(* Logix 5000 project; controller CIP_14485201 vendor 1 type 14 code 216 rev 38.11; software revision 38.01; part 10 of 11 *)
(* tags used below, declared in another part *)
   Bit : BOOL[128];   // BIT
   CIP_to_Process : CIP_to_Process;   // CIP TO PROCESS SIGNALS
   cipToProcess : BOOL;   // send signal to dcs
   Heartbeat_to_dcs_off : TIMER;   // 5 second toggle
   heartbeat_to_dcs_on : TIMER;   // turns on heartbeat to dcs
   Messages_List : STRING;   // ACTIVE MESSAGES ECHO FROM HMI
   MOA_Drain_Flow_Mod_Value : INT;   // PV MOA DRAIN FLOW MODULATION VALUE
   MOA_Drain_Flow_Mod_Value_Status : BOOL;   // PV MOA DRAIN FLOW MODULATION VALUE STATUS BIT
   MOA_OFF : DINT[20];   // PANELVIEW MOA OFF
   MOA_ON : DINT[20];   // PANELVIEW MOA ON
   Opcode_Description : STRING;   // ACTIVE OPCODE ECHO FROM HMI
   OpCode_Pin : DINT[5];   // OPCODE PIN ARRAY
   Panelview : INT[40];   // PANELVIEW CONTROL
   PID2 : PID;   // SUPPLY FLOW PID
   Process_Heartbeat_Memory : BOOL;
   Process_to_CIP : Process_to_CIP;   // PROCESS SIGNALS TO CIP
   pv_step_time_minutes : DINT;   // PANELVIEW DISPLAY STEP TIME MINUTES
   pv_step_time_seconds : DINT;   // PANELVIEW DISPLAY STEP TIME SECONDS
   Recipe : RECIPE[41];   // RECIPES
   SCLD_Drain_Flow : SCALE;   // DRAIN FLOW MODULATION 0-100%
   SCLD_DrainValve_Feedback : SCALE;   // DRAIN FLOW FEEDBACK POSITION 0-100%
   SCLD_Return_Temp : SCALE;   // RETURN TEMPERATURE 0-100°C
   SCLD_Rinse_Cond : SCALE;   // RINSE CONDUCTIVITY 0-10 uS/cm
   SCLD_Supply_Flow : SCALE;   // SUPPLY FLOW 0-60 GPM
   SCLD_Supply_Press : SCALE;   // SUPPLY PRESSURE 0-100 PSIG
   SCLD_Supply_Temp : SCALE;   // SUPPLY TEMPERATURE 0-100°C
   SCLD_SupplyValve_Feedback : SCALE;   // SUPPLY FLOW FEEDBACK POSITION 0-100%
   SCLD_Wash_Cond : SCALE;   // WASH CONDUCTIVITY 0-100 mS/cm
   Sequencer : CONTROL[4];   // SEQUENCER
   SP_Drain_Flow : REAL;   // CURRENT DRAIN FLOW MODULATION SETPOINT
   SP_DrainValve_HighDeadband : REAL;   // CURRENT DRAIN VALVE DEADBAND SETPOINT
   SP_DrainValve_LowDeadband : REAL;   // CURRENT DRAIN VALVE DEADBAND SETPOINT
   SP_Supply_Flow : REAL;   // CURRENT SUPPLY FLOW SETPOINT
   SP_SupplyValve_HighDeadband : REAL;   // CURRENT SUPPLY VALVE DEADBAND SETPOINT
   SP_SupplyValve_LowDeadband : REAL;   // CURRENT SUPPLY VALVE DEADBAND SETPOINT
   Step_Time_Min : STRING;
   Step_Time_Remaining : STRING[5];
   Step_Time_Sec : STRING;
   Timer : TIMER[99];   // TIMER
   Timer_Chem1_Pump : TIMER[7];   // CHEM #1 CONTROL TIMERS
   Timer_Chem2_Pump : TIMER[7];   // CHEM #2 CONTROL TIMERS
   Utility_Out : DINT[5];   // PANELVIEW UTILITY OUTPUT CONTROL
(* MainProgram, continued *)

ROUTINE _88_LEVEL   (* ladder *)
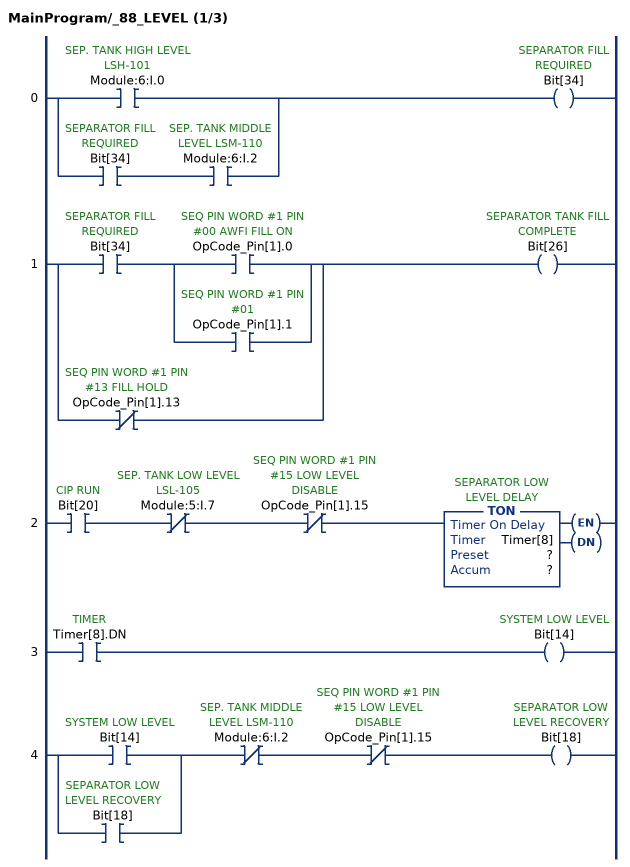
   0: [XIC(Module:6:I.0) ,XIC(Bit[34]) XIC(Module:6:I.2) ]OTE(Bit[34]);
   1: [XIC(Bit[34]) [XIC(OpCode_Pin[1].0) ,XIC(OpCode_Pin[1].1) ] ,XIO(OpCode_Pin[1].13) ]OTE(Bit[26]);
   2: XIC(Bit[20])XIO(Module:5:I.7)XIO(OpCode_Pin[1].15)TON(Timer[8],?,?);
   3: XIC(Timer[8].DN)OTE(Bit[14]);
   4: [XIC(Bit[14]) ,XIC(Bit[18]) ]XIO(Module:6:I.2)XIO(OpCode_Pin[1].15)OTE(Bit[18]);
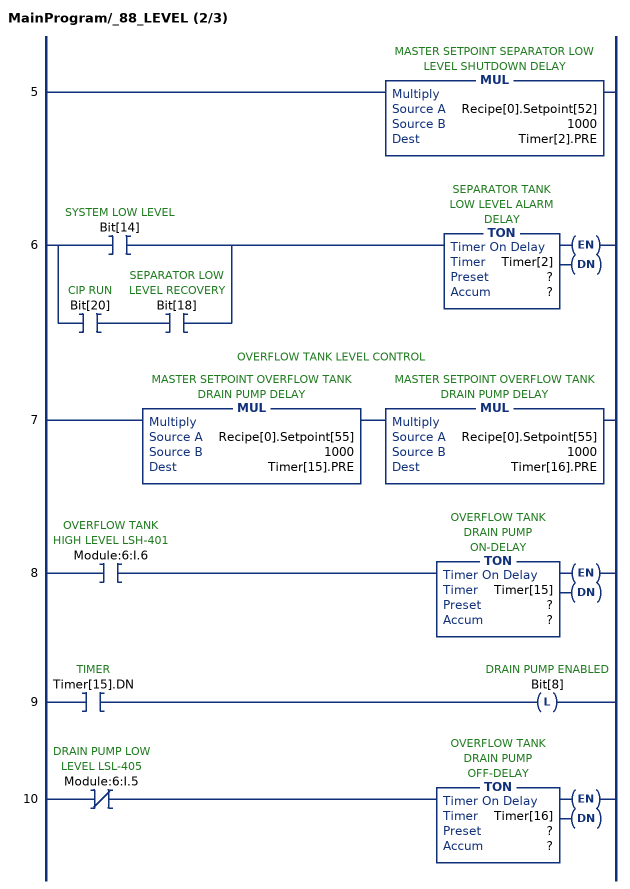
   5: MUL(Recipe[0].Setpoint[52],1000,Timer[2].PRE);
   6: [XIC(Bit[14]) ,XIC(Bit[20]) XIC(Bit[18]) ]TON(Timer[2],?,?);
   // OVERFLOW TANK LEVEL CONTROL
   7: MUL(Recipe[0].Setpoint[55],1000,Timer[15].PRE)MUL(Recipe[0].Setpoint[55],1000,Timer[16].PRE);
   8: XIC(Module:6:I.6)TON(Timer[15],?,?);
   9: XIC(Timer[15].DN)OTL(Bit[8]);
   10: XIO(Module:6:I.5)TON(Timer[16],?,?);
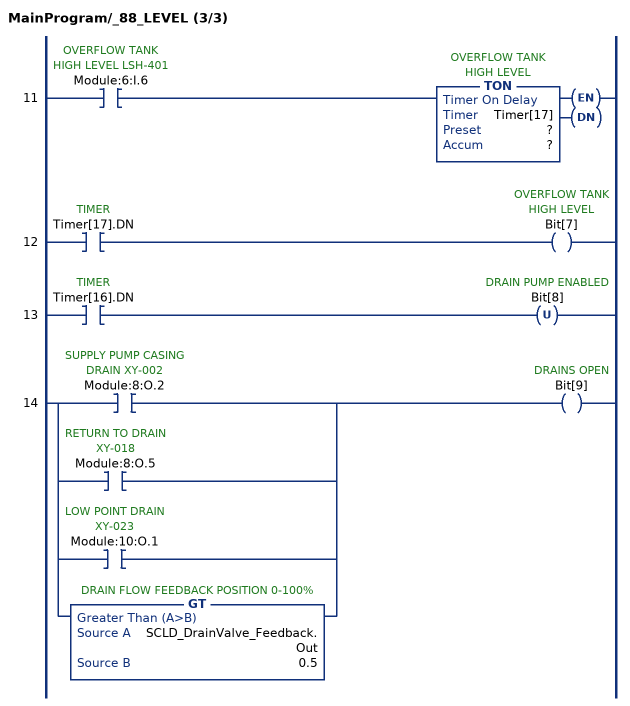
   11: XIC(Module:6:I.6)TON(Timer[17],?,?);
   12: XIC(Timer[17].DN)OTE(Bit[7]);
   13: XIC(Timer[16].DN)OTU(Bit[8]);
   14: [XIC(Module:8:O.2) ,XIC(Module:8:O.5) ,XIC(Module:10:O.1) ,GT(SCLD_DrainValve_Feedback.Out,0.5) ]OTE(Bit[9]);
END_ROUTINE

ROUTINE _89_FLOW   (* ladder *)
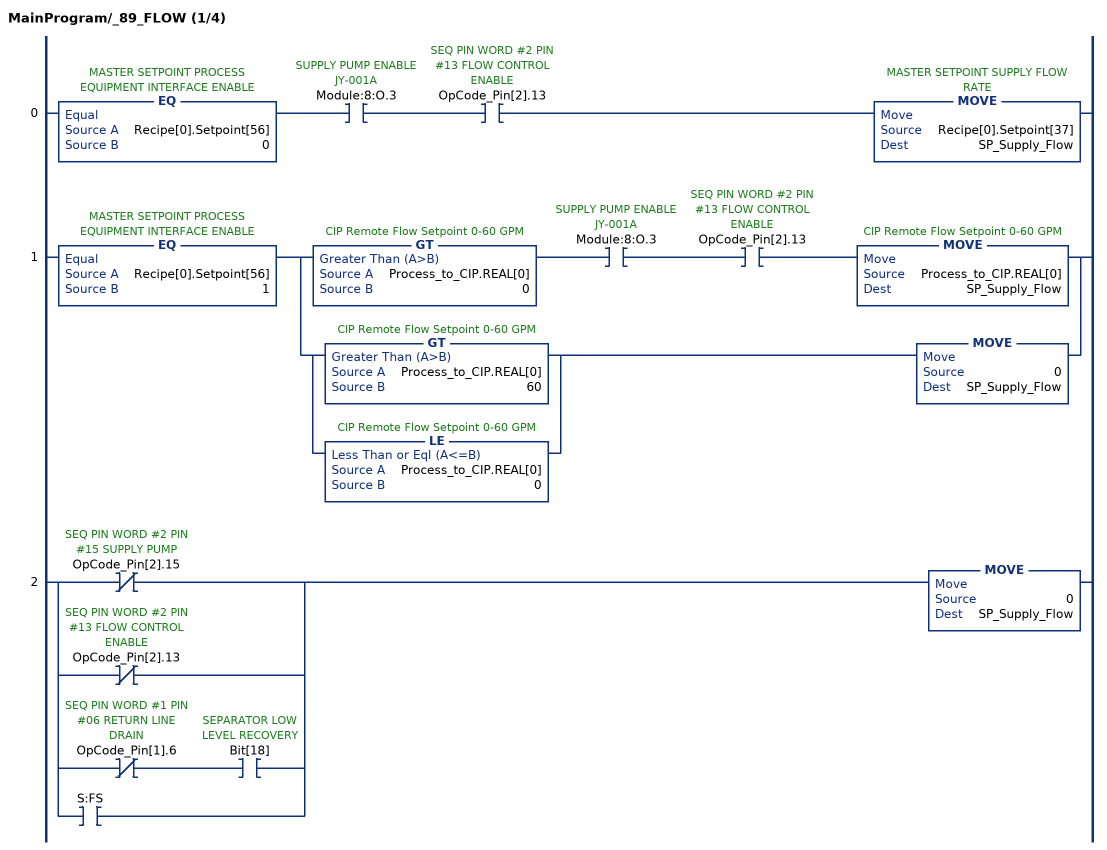
   0: EQ(Recipe[0].Setpoint[56],0)XIC(Module:8:O.3)XIC(OpCode_Pin[2].13)MOVE(Recipe[0].Setpoint[37],SP_Supply_Flow);
   1: EQ(Recipe[0].Setpoint[56],1)[GT(Process_to_CIP.REAL[0],0) XIC(Module:8:O.3) XIC(OpCode_Pin[2].13) MOVE(Process_to_CIP.REAL[0],SP_Supply_Flow) ,[GT(Process_to_CIP.REAL[0],60) ,LE(Process_to_CIP.REAL[0],0) ] MOVE(0,SP_Supply_Flow) ];
   2: [XIO(OpCode_Pin[2].15) ,XIO(OpCode_Pin[2].13) ,XIO(OpCode_Pin[1].6) XIC(Bit[18]) ,XIC(S:FS) ]MOVE(0,SP_Supply_Flow);
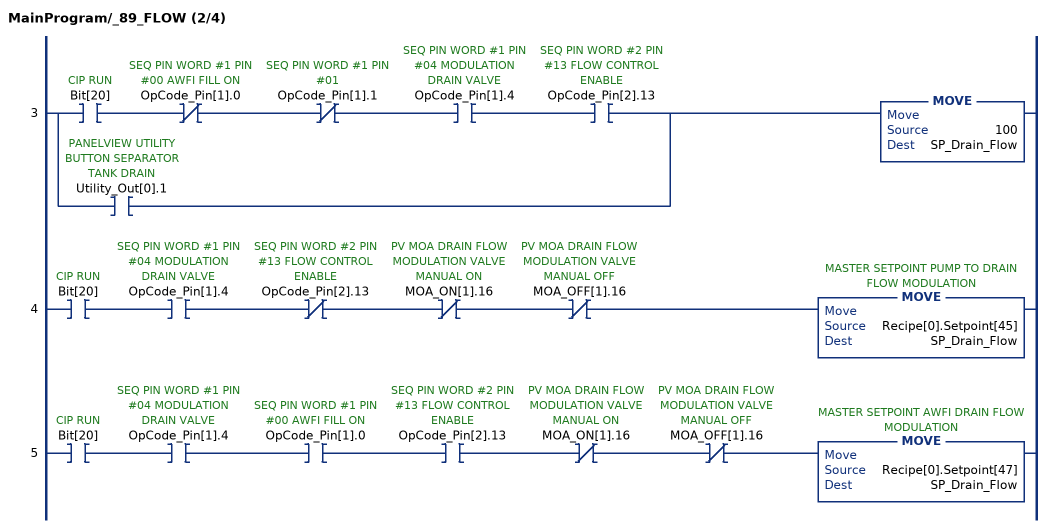
   3: [XIC(Bit[20]) XIO(OpCode_Pin[1].0) XIO(OpCode_Pin[1].1) XIC(OpCode_Pin[1].4) XIC(OpCode_Pin[2].13) ,XIC(Utility_Out[0].1) ]MOVE(100,SP_Drain_Flow);
   4: XIC(Bit[20])XIC(OpCode_Pin[1].4)XIO(OpCode_Pin[2].13)XIO(MOA_ON[1].16)XIO(MOA_OFF[1].16)MOVE(Recipe[0].Setpoint[45],SP_Drain_Flow);
   5: XIC(Bit[20])XIC(OpCode_Pin[1].4)XIC(OpCode_Pin[1].0)XIC(OpCode_Pin[2].13)XIO(MOA_ON[1].16)XIO(MOA_OFF[1].16)MOVE(Recipe[0].Setpoint[47],SP_Drain_Flow);
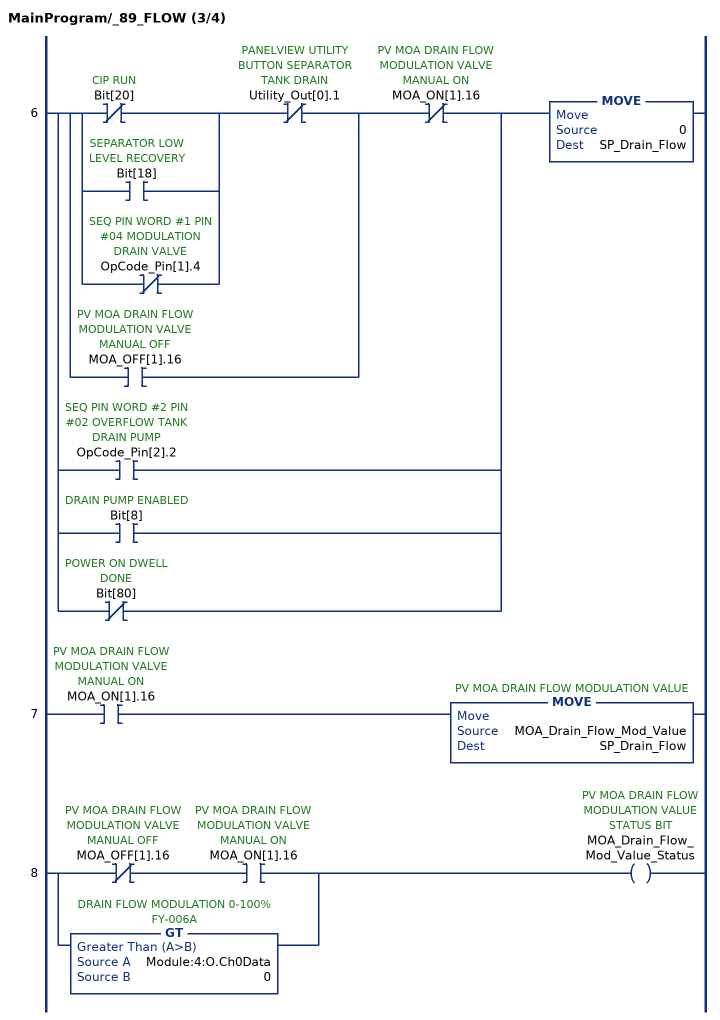
   6: [[[XIO(Bit[20]) ,XIC(Bit[18]) ,XIO(OpCode_Pin[1].4) ] XIO(Utility_Out[0].1) ,XIC(MOA_OFF[1].16) ] XIO(MOA_ON[1].16) ,XIC(OpCode_Pin[2].2) ,XIC(Bit[8]) ,XIO(Bit[80]) ]MOVE(0,SP_Drain_Flow);
   7: XIC(MOA_ON[1].16)MOVE(MOA_Drain_Flow_Mod_Value,SP_Drain_Flow);
   8: [XIO(MOA_OFF[1].16) XIC(MOA_ON[1].16) ,GT(Module:4:O.Ch0Data,0) ]OTE(MOA_Drain_Flow_Mod_Value_Status);
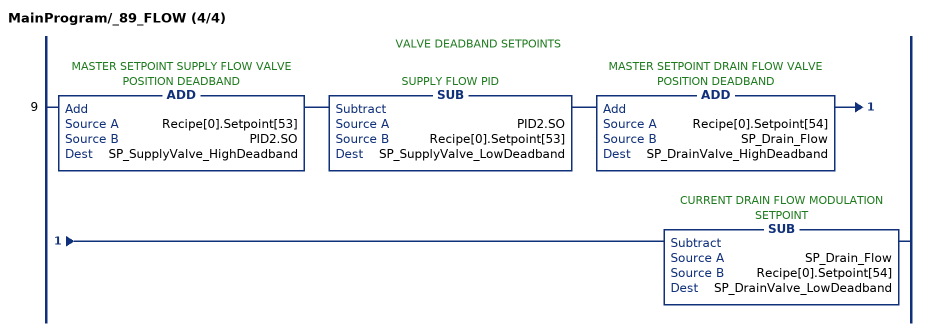
   // VALVE DEADBAND SETPOINTS
   9: ADD(Recipe[0].Setpoint[53],PID2.SO,SP_SupplyValve_HighDeadband)SUB(PID2.SO,Recipe[0].Setpoint[53],SP_SupplyValve_LowDeadband)ADD(Recipe[0].Setpoint[54],SP_Drain_Flow,SP_DrainValve_HighDeadband)SUB(SP_Drain_Flow,Recipe[0].Setpoint[54],SP_DrainValve_LowDeadband);
END_ROUTINE

ROUTINE _90_OUTPUTS   (* ladder *)
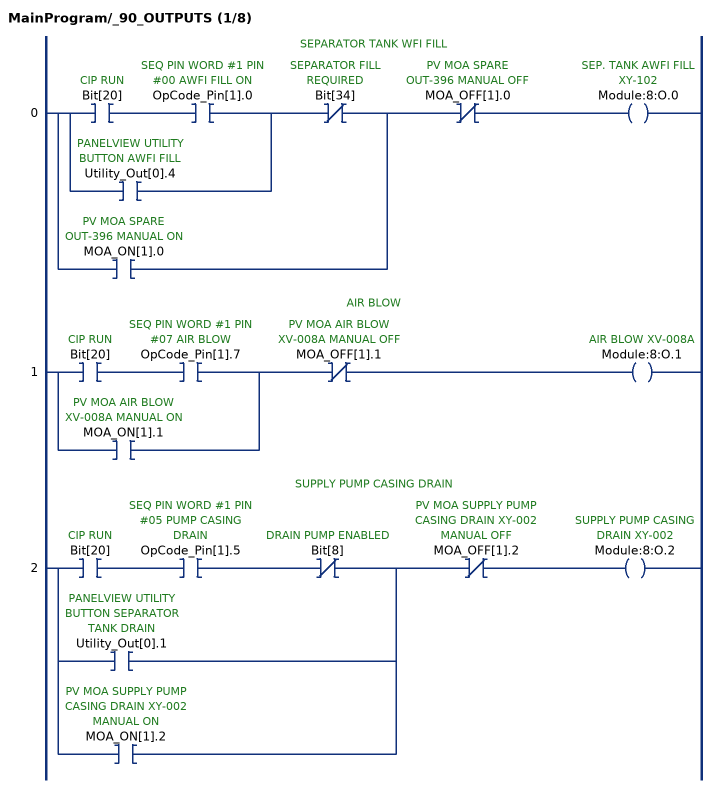
   // SEPARATOR TANK WFI FILL
   0: [[XIC(Bit[20]) XIC(OpCode_Pin[1].0) ,XIC(Utility_Out[0].4) ] XIO(Bit[34]) ,XIC(MOA_ON[1].0) ]XIO(MOA_OFF[1].0)OTE(Module:8:O.0);
   // AIR BLOW
   1: [XIC(Bit[20]) XIC(OpCode_Pin[1].7) ,XIC(MOA_ON[1].1) ]XIO(MOA_OFF[1].1)OTE(Module:8:O.1);
   // SUPPLY PUMP CASING DRAIN
   2: [XIC(Bit[20]) XIC(OpCode_Pin[1].5) XIO(Bit[8]) ,XIC(Utility_Out[0].1) ,XIC(MOA_ON[1].2) ]XIO(MOA_OFF[1].2)OTE(Module:8:O.2);
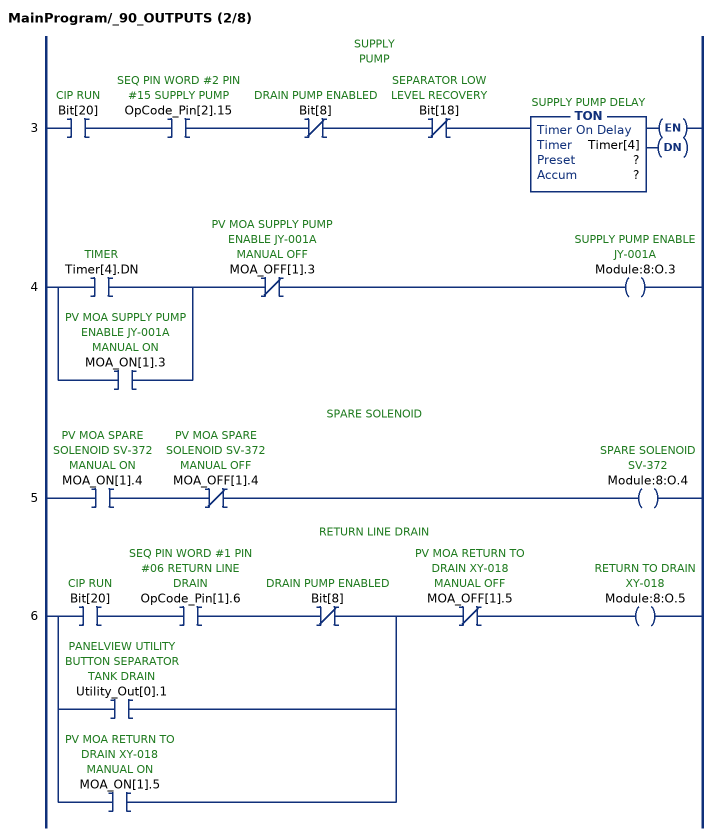
   // SUPPLY
   // PUMP
   3: XIC(Bit[20])XIC(OpCode_Pin[2].15)XIO(Bit[8])XIO(Bit[18])TON(Timer[4],?,?);
   4: [XIC(Timer[4].DN) ,XIC(MOA_ON[1].3) ]XIO(MOA_OFF[1].3)OTE(Module:8:O.3);
   // SPARE SOLENOID
   5: XIC(MOA_ON[1].4)XIO(MOA_OFF[1].4)OTE(Module:8:O.4);
   // RETURN LINE DRAIN
   6: [XIC(Bit[20]) XIC(OpCode_Pin[1].6) XIO(Bit[8]) ,XIC(Utility_Out[0].1) ,XIC(MOA_ON[1].5) ]XIO(MOA_OFF[1].5)OTE(Module:8:O.5);
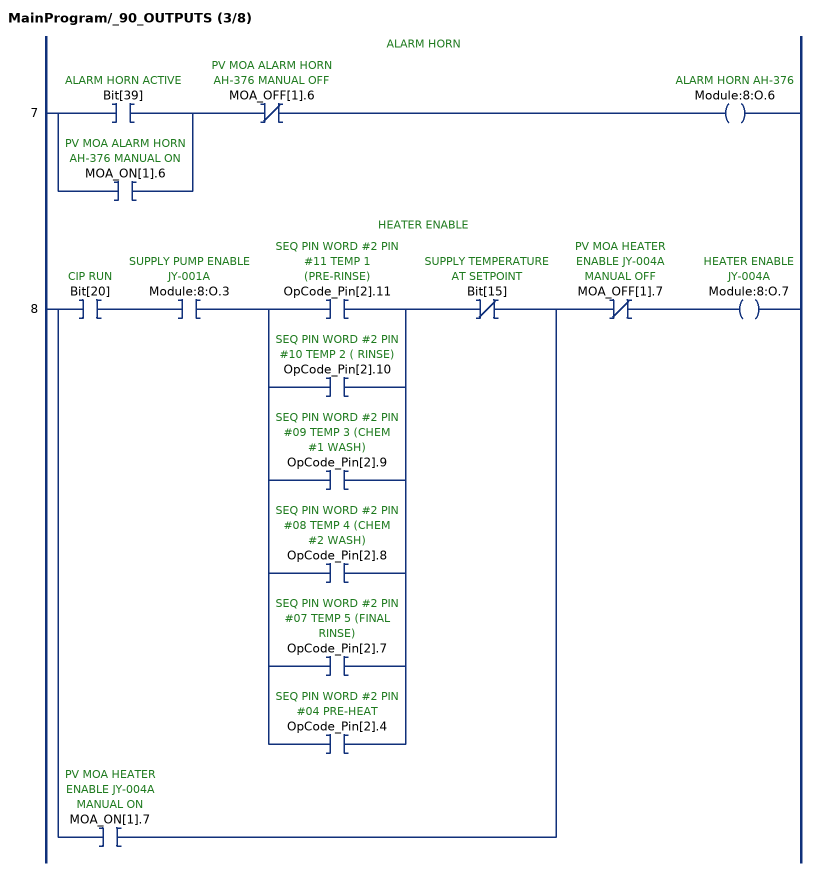
   // ALARM HORN
   7: [XIC(Bit[39]) ,XIC(MOA_ON[1].6) ]XIO(MOA_OFF[1].6)OTE(Module:8:O.6);
   // HEATER ENABLE
   8: [XIC(Bit[20]) XIC(Module:8:O.3) [XIC(OpCode_Pin[2].11) ,XIC(OpCode_Pin[2].10) ,XIC(OpCode_Pin[2].9) ,XIC(OpCode_Pin[2].8) ,XIC(OpCode_Pin[2].7) ,XIC(OpCode_Pin[2].4) ] XIO(Bit[15]) ,XIC(MOA_ON[1].7) ]XIO(MOA_OFF[1].7)OTE(Module:8:O.7);
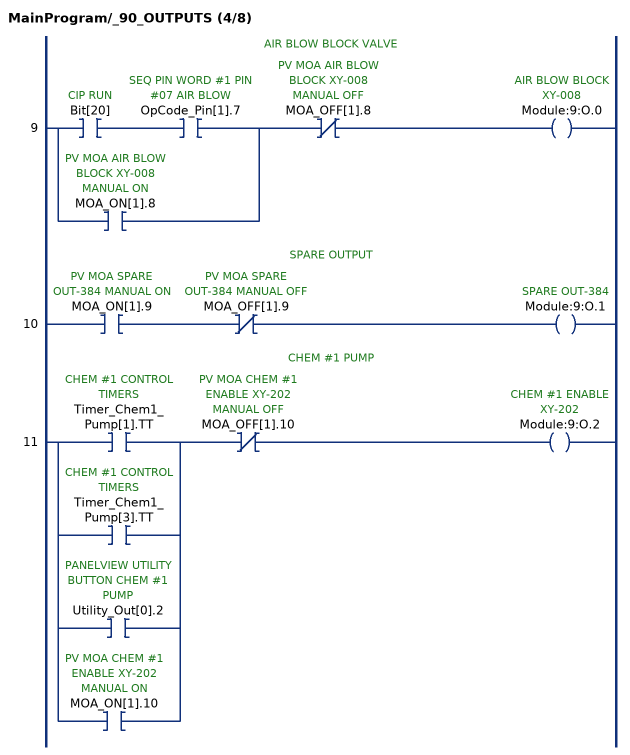
   // AIR BLOW BLOCK VALVE
   9: [XIC(Bit[20]) XIC(OpCode_Pin[1].7) ,XIC(MOA_ON[1].8) ]XIO(MOA_OFF[1].8)OTE(Module:9:O.0);
   // SPARE OUTPUT
   10: XIC(MOA_ON[1].9)XIO(MOA_OFF[1].9)OTE(Module:9:O.1);
   // CHEM #1 PUMP
   11: [XIC(Timer_Chem1_Pump[1].TT) ,XIC(Timer_Chem1_Pump[3].TT) ,XIC(Utility_Out[0].2) ,XIC(MOA_ON[1].10) ]XIO(MOA_OFF[1].10)OTE(Module:9:O.2);
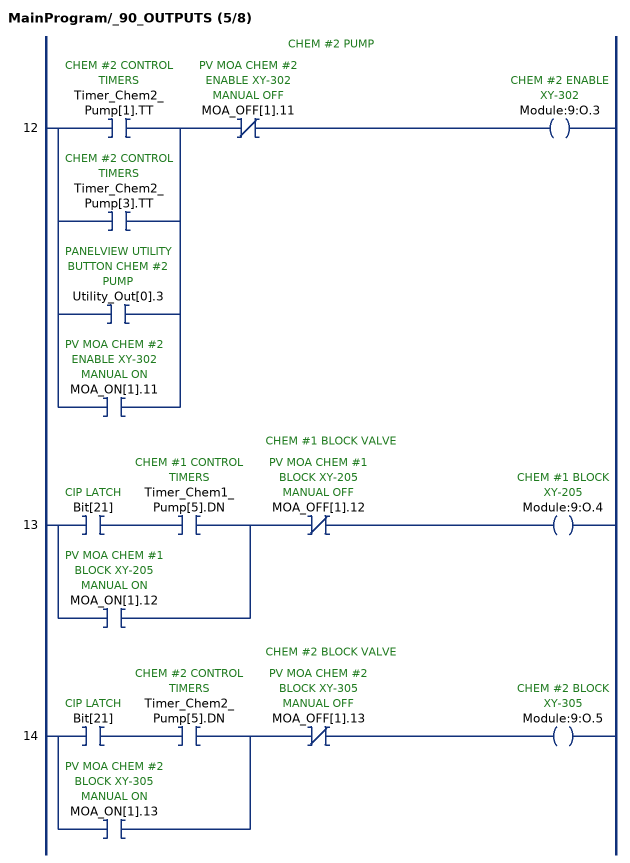
   // CHEM #2 PUMP
   12: [XIC(Timer_Chem2_Pump[1].TT) ,XIC(Timer_Chem2_Pump[3].TT) ,XIC(Utility_Out[0].3) ,XIC(MOA_ON[1].11) ]XIO(MOA_OFF[1].11)OTE(Module:9:O.3);
   // CHEM #1 BLOCK VALVE
   13: [XIC(Bit[21]) XIC(Timer_Chem1_Pump[5].DN) ,XIC(MOA_ON[1].12) ]XIO(MOA_OFF[1].12)OTE(Module:9:O.4);
   // CHEM #2 BLOCK VALVE
   14: [XIC(Bit[21]) XIC(Timer_Chem2_Pump[5].DN) ,XIC(MOA_ON[1].13) ]XIO(MOA_OFF[1].13)OTE(Module:9:O.5);
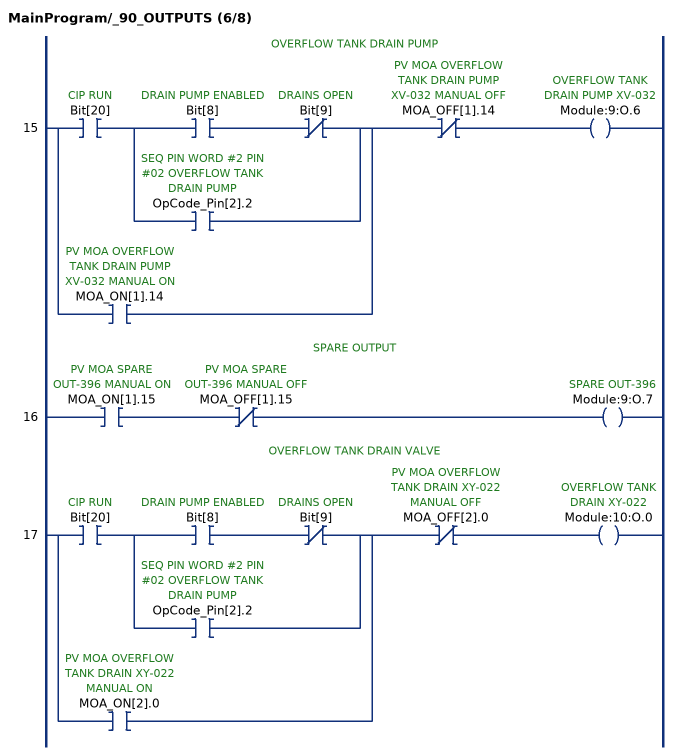
   // OVERFLOW TANK DRAIN PUMP
   15: [XIC(Bit[20]) [XIC(Bit[8]) XIO(Bit[9]) ,XIC(OpCode_Pin[2].2) ] ,XIC(MOA_ON[1].14) ]XIO(MOA_OFF[1].14)OTE(Module:9:O.6);
   // SPARE OUTPUT
   16: XIC(MOA_ON[1].15)XIO(MOA_OFF[1].15)OTE(Module:9:O.7);
   // OVERFLOW TANK DRAIN VALVE
   17: [XIC(Bit[20]) [XIC(Bit[8]) XIO(Bit[9]) ,XIC(OpCode_Pin[2].2) ] ,XIC(MOA_ON[2].0) ]XIO(MOA_OFF[2].0)OTE(Module:10:O.0);
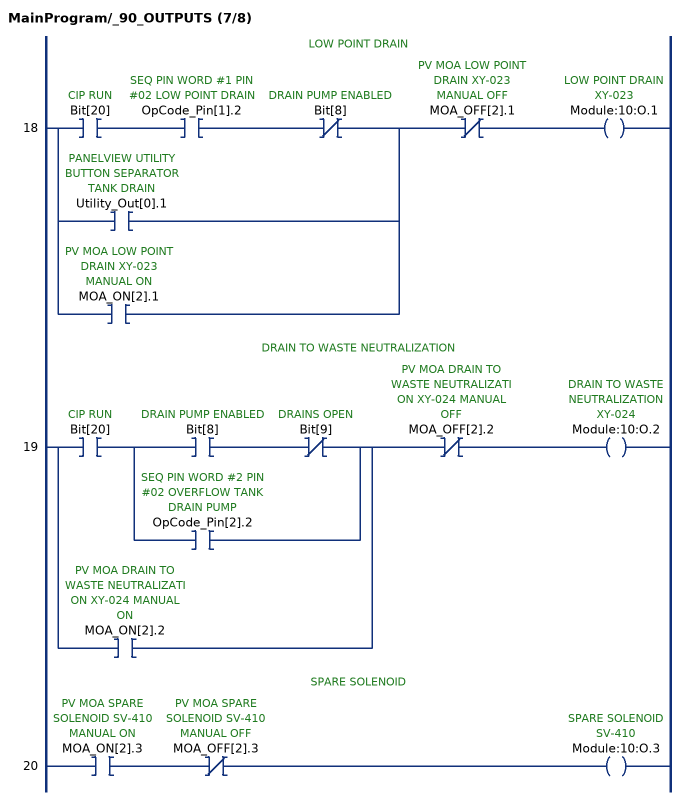
   // LOW POINT DRAIN
   18: [XIC(Bit[20]) XIC(OpCode_Pin[1].2) XIO(Bit[8]) ,XIC(Utility_Out[0].1) ,XIC(MOA_ON[2].1) ]XIO(MOA_OFF[2].1)OTE(Module:10:O.1);
   // DRAIN TO WASTE NEUTRALIZATION
   19: [XIC(Bit[20]) [XIC(Bit[8]) XIO(Bit[9]) ,XIC(OpCode_Pin[2].2) ] ,XIC(MOA_ON[2].2) ]XIO(MOA_OFF[2].2)OTE(Module:10:O.2);
   // SPARE SOLENOID
   20: XIC(MOA_ON[2].3)XIO(MOA_OFF[2].3)OTE(Module:10:O.3);
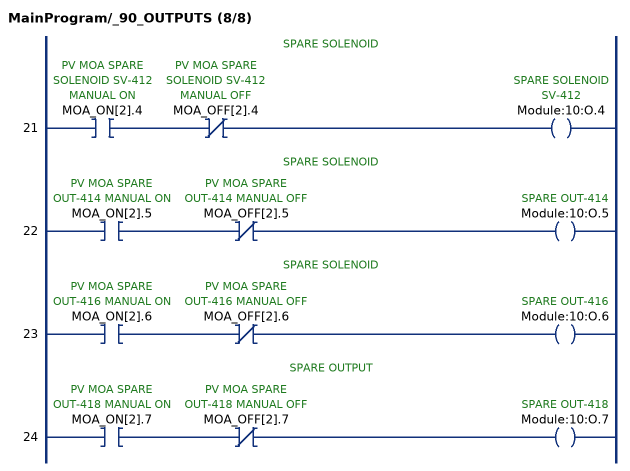
   // SPARE SOLENOID
   21: XIC(MOA_ON[2].4)XIO(MOA_OFF[2].4)OTE(Module:10:O.4);
   // SPARE SOLENOID
   22: XIC(MOA_ON[2].5)XIO(MOA_OFF[2].5)OTE(Module:10:O.5);
   // SPARE SOLENOID
   23: XIC(MOA_ON[2].6)XIO(MOA_OFF[2].6)OTE(Module:10:O.6);
   // SPARE OUTPUT
   24: XIC(MOA_ON[2].7)XIO(MOA_OFF[2].7)OTE(Module:10:O.7);
END_ROUTINE

ROUTINE _99_COMMS   (* ladder *)
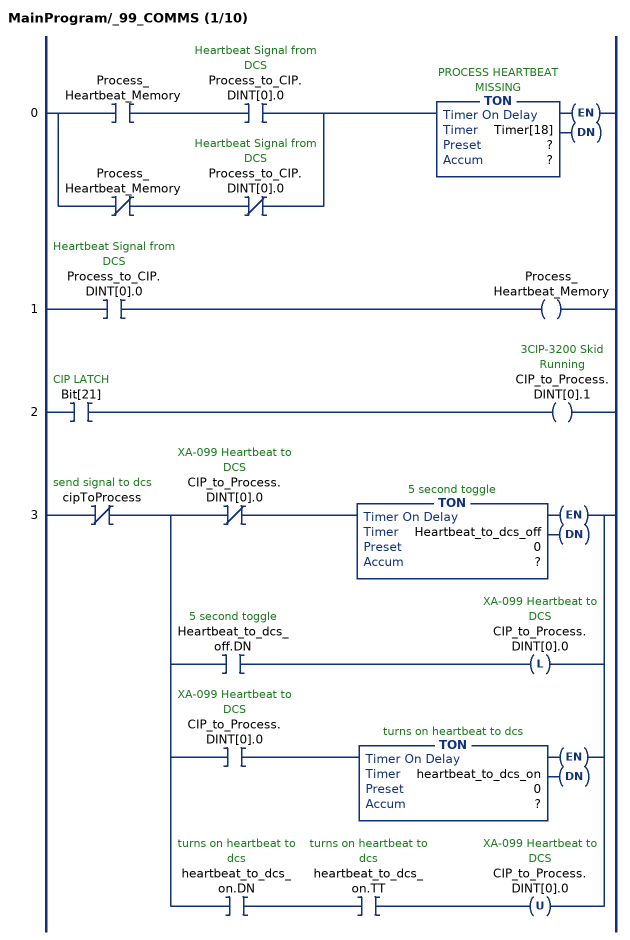
   0: [XIC(Process_Heartbeat_Memory) XIC(Process_to_CIP.DINT[0].0) ,XIO(Process_Heartbeat_Memory) XIO(Process_to_CIP.DINT[0].0) ]TON(Timer[18],?,?);
   1: XIC(Process_to_CIP.DINT[0].0)OTE(Process_Heartbeat_Memory);
   2: XIC(Bit[21])OTE(CIP_to_Process.DINT[0].1);
   3: XIO(cipToProcess)[XIO(CIP_to_Process.DINT[0].0) TON(Heartbeat_to_dcs_off,?,?) ,XIC(Heartbeat_to_dcs_off.DN) OTL(CIP_to_Process.DINT[0].0) ,XIC(CIP_to_Process.DINT[0].0) TON(heartbeat_to_dcs_on,?,?) ,XIC(heartbeat_to_dcs_on.DN) XIC(heartbeat_to_dcs_on.TT) OTU(CIP_to_Process.DINT[0].0) ];
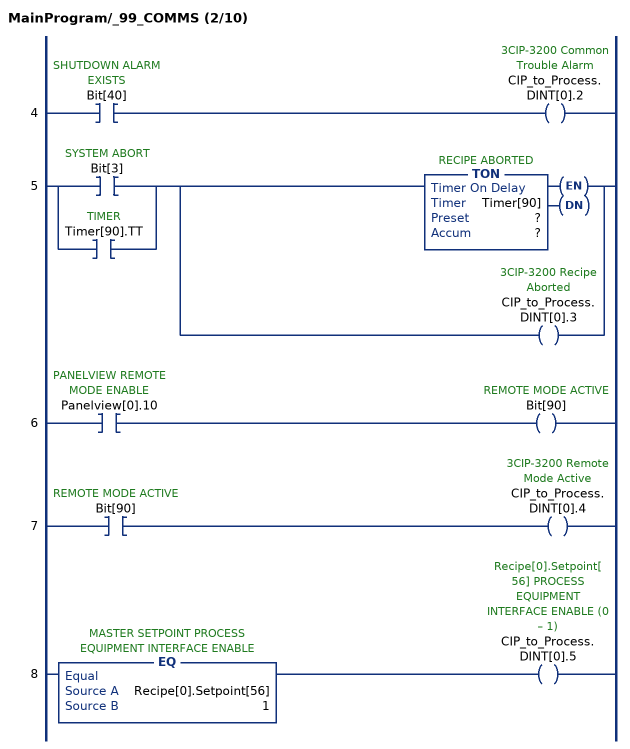
   4: XIC(Bit[40])OTE(CIP_to_Process.DINT[0].2);
   5: [XIC(Bit[3]) ,XIC(Timer[90].TT) ][TON(Timer[90],?,?) ,OTE(CIP_to_Process.DINT[0].3) ];
   6: XIC(Panelview[0].10)OTE(Bit[90]);
   7: XIC(Bit[90])OTE(CIP_to_Process.DINT[0].4);
   8: EQ(Recipe[0].Setpoint[56],1)OTE(CIP_to_Process.DINT[0].5);
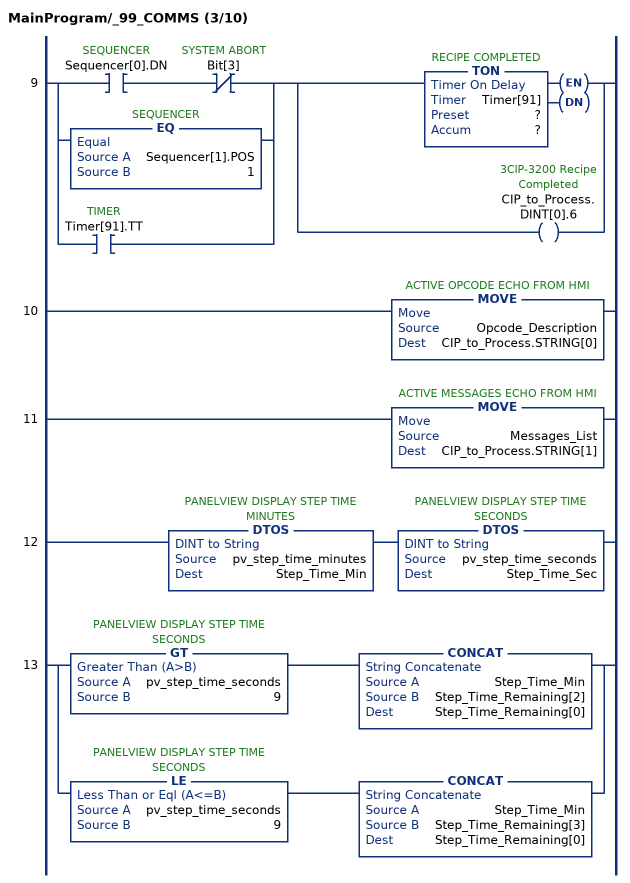
   9: [XIC(Sequencer[0].DN) XIO(Bit[3]) ,EQ(Sequencer[1].POS,1) ,XIC(Timer[91].TT) ][TON(Timer[91],?,?) ,OTE(CIP_to_Process.DINT[0].6) ];
   10: MOVE(Opcode_Description,CIP_to_Process.STRING[0]);
   11: MOVE(Messages_List,CIP_to_Process.STRING[1]);
   12: DTOS(pv_step_time_minutes,Step_Time_Min)DTOS(pv_step_time_seconds,Step_Time_Sec);
   13: [GT(pv_step_time_seconds,9) CONCAT(Step_Time_Min,Step_Time_Remaining[2],Step_Time_Remaining[0]) ,LE(pv_step_time_seconds,9) CONCAT(Step_Time_Min,Step_Time_Remaining[3],Step_Time_Remaining[0]) ];
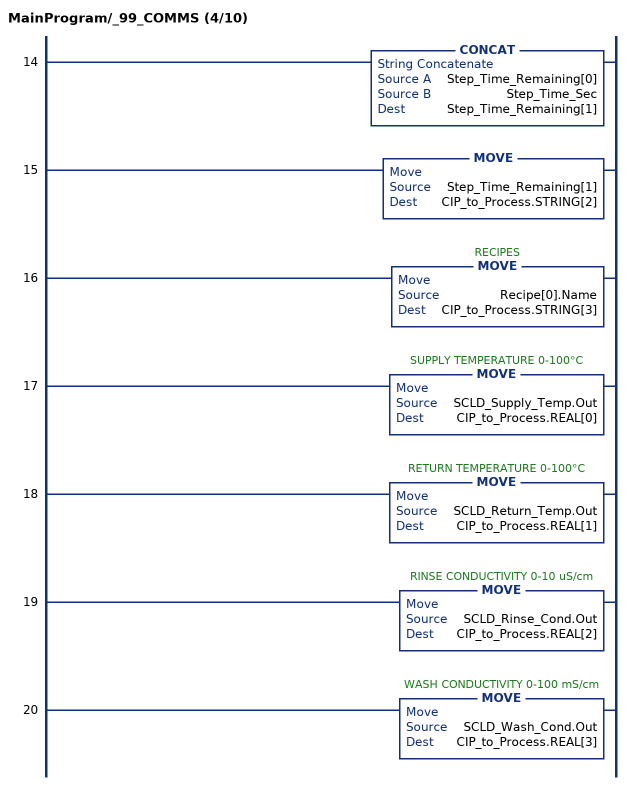
   14: CONCAT(Step_Time_Remaining[0],Step_Time_Sec,Step_Time_Remaining[1]);
   15: MOVE(Step_Time_Remaining[1],CIP_to_Process.STRING[2]);
   16: MOVE(Recipe[0].Name,CIP_to_Process.STRING[3]);
   17: MOVE(SCLD_Supply_Temp.Out,CIP_to_Process.REAL[0]);
   18: MOVE(SCLD_Return_Temp.Out,CIP_to_Process.REAL[1]);
   19: MOVE(SCLD_Rinse_Cond.Out,CIP_to_Process.REAL[2]);
   20: MOVE(SCLD_Wash_Cond.Out,CIP_to_Process.REAL[3]);
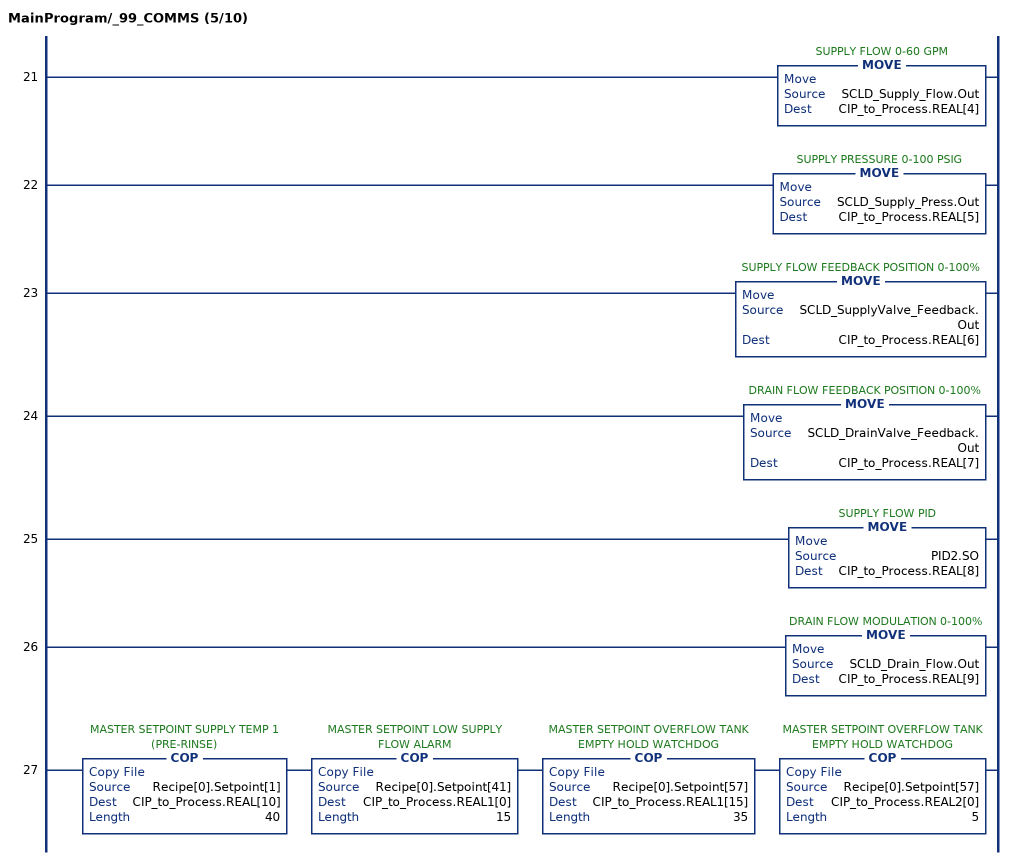
   21: MOVE(SCLD_Supply_Flow.Out,CIP_to_Process.REAL[4]);
   22: MOVE(SCLD_Supply_Press.Out,CIP_to_Process.REAL[5]);
   23: MOVE(SCLD_SupplyValve_Feedback.Out,CIP_to_Process.REAL[6]);
   24: MOVE(SCLD_DrainValve_Feedback.Out,CIP_to_Process.REAL[7]);
   25: MOVE(PID2.SO,CIP_to_Process.REAL[8]);
   26: MOVE(SCLD_Drain_Flow.Out,CIP_to_Process.REAL[9]);
   27: COP(Recipe[0].Setpoint[1],CIP_to_Process.REAL[10],40)COP(Recipe[0].Setpoint[41],CIP_to_Process.REAL1[0],15)COP(Recipe[0].Setpoint[57],CIP_to_Process.REAL1[15],35)COP(Recipe[0].Setpoint[57],CIP_to_Process.REAL2[0],5);
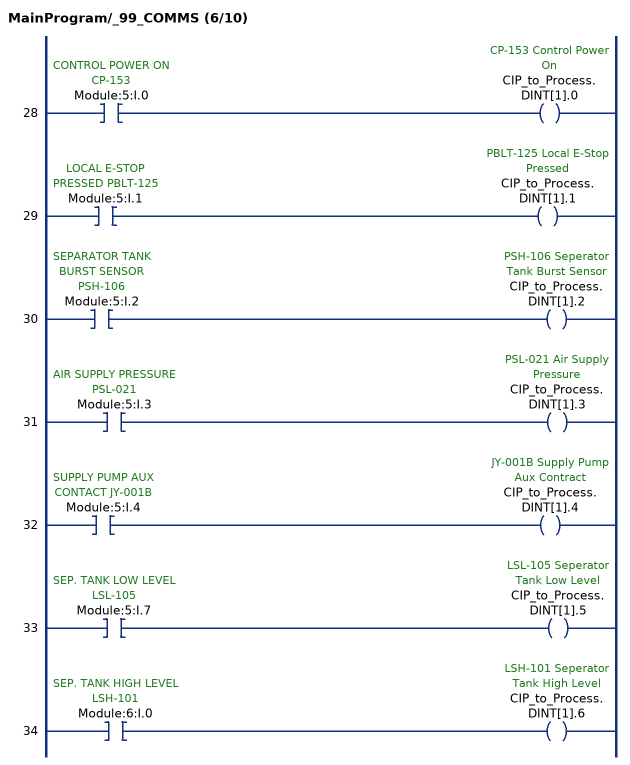
   28: XIC(Module:5:I.0)OTE(CIP_to_Process.DINT[1].0);
   29: XIC(Module:5:I.1)OTE(CIP_to_Process.DINT[1].1);
   30: XIC(Module:5:I.2)OTE(CIP_to_Process.DINT[1].2);
   31: XIC(Module:5:I.3)OTE(CIP_to_Process.DINT[1].3);
   32: XIC(Module:5:I.4)OTE(CIP_to_Process.DINT[1].4);
   33: XIC(Module:5:I.7)OTE(CIP_to_Process.DINT[1].5);
   34: XIC(Module:6:I.0)OTE(CIP_to_Process.DINT[1].6);
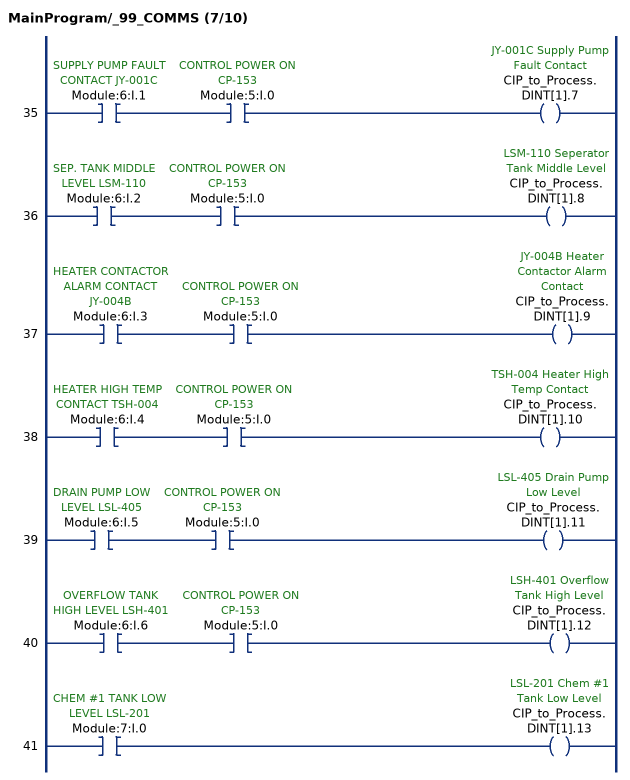
   35: XIC(Module:6:I.1)XIC(Module:5:I.0)OTE(CIP_to_Process.DINT[1].7);
   36: XIC(Module:6:I.2)XIC(Module:5:I.0)OTE(CIP_to_Process.DINT[1].8);
   37: XIC(Module:6:I.3)XIC(Module:5:I.0)OTE(CIP_to_Process.DINT[1].9);
   38: XIC(Module:6:I.4)XIC(Module:5:I.0)OTE(CIP_to_Process.DINT[1].10);
   39: XIC(Module:6:I.5)XIC(Module:5:I.0)OTE(CIP_to_Process.DINT[1].11);
   40: XIC(Module:6:I.6)XIC(Module:5:I.0)OTE(CIP_to_Process.DINT[1].12);
   41: XIC(Module:7:I.0)OTE(CIP_to_Process.DINT[1].13);
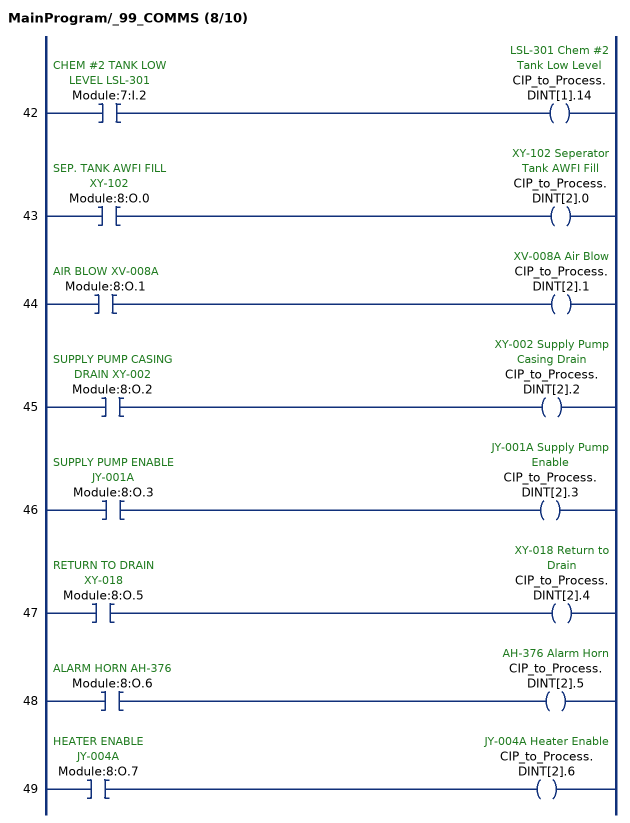
   42: XIC(Module:7:I.2)OTE(CIP_to_Process.DINT[1].14);
   43: XIC(Module:8:O.0)OTE(CIP_to_Process.DINT[2].0);
   44: XIC(Module:8:O.1)OTE(CIP_to_Process.DINT[2].1);
   45: XIC(Module:8:O.2)OTE(CIP_to_Process.DINT[2].2);
   46: XIC(Module:8:O.3)OTE(CIP_to_Process.DINT[2].3);
   47: XIC(Module:8:O.5)OTE(CIP_to_Process.DINT[2].4);
   48: XIC(Module:8:O.6)OTE(CIP_to_Process.DINT[2].5);
   49: XIC(Module:8:O.7)OTE(CIP_to_Process.DINT[2].6);
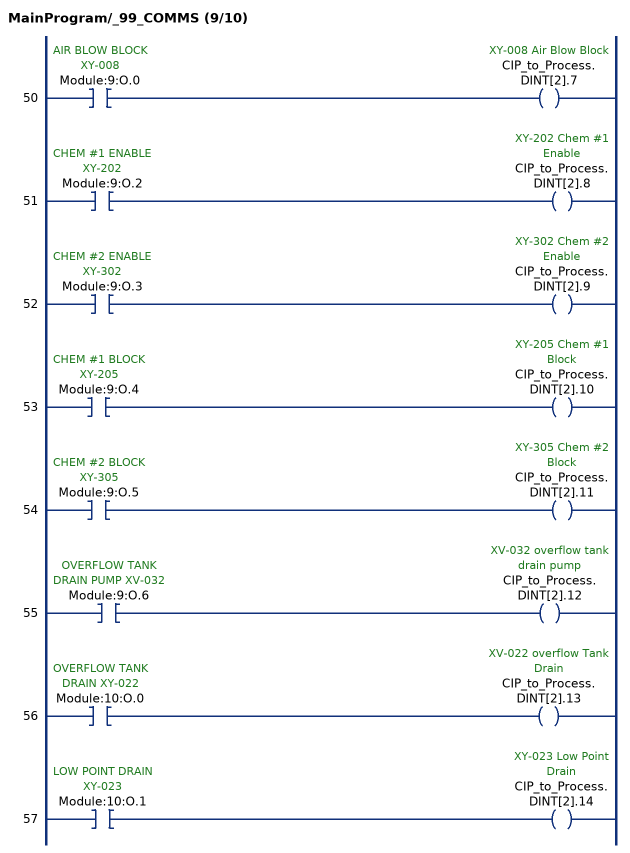
   50: XIC(Module:9:O.0)OTE(CIP_to_Process.DINT[2].7);
   51: XIC(Module:9:O.2)OTE(CIP_to_Process.DINT[2].8);
   52: XIC(Module:9:O.3)OTE(CIP_to_Process.DINT[2].9);
   53: XIC(Module:9:O.4)OTE(CIP_to_Process.DINT[2].10);
   54: XIC(Module:9:O.5)OTE(CIP_to_Process.DINT[2].11);
   55: XIC(Module:9:O.6)OTE(CIP_to_Process.DINT[2].12);
   56: XIC(Module:10:O.0)OTE(CIP_to_Process.DINT[2].13);
   57: XIC(Module:10:O.1)OTE(CIP_to_Process.DINT[2].14);
